// TIA Portal V21 export
// export: Created 2026-11-22T02:34:22.6112688Z, ExportSetting WithDefaults, DisplayName Totally Integrated Automation Portal, DisplayVersion V21 Update 3, DisplayName STEP 7 Professional, DisplayVersion V21 Update 3, DisplayName STEP 7 Safety, DisplayVersion V21, DisplayName Tech WebApplication, DisplayVersion V21, DisplayName WinCC Basic/Comfort/Advanced, DisplayVersion V21 Update 3, DisplayName WinCC Unified, DisplayVersion V21 Update 3
TextList "TL_Value"  ListRange=Decimal
  TextListEntry   EntryType=Range, From=-100, To=-1, Text="Negative (-100..-1)"
  TextListEntry   EntryType=SingleValue, Text="Zero"
  TextListEntry   EntryType=Range, From=1, To=9, Text="One to nine"
  TextListEntry   EntryType=SingleValue, From=10, To=10, Text="Ten: Ünïcödé äöüß ÄÖÜ €"
  TextListEntry   EntryType=SingleValue, From=32000, To=32000, Text="Undefined value (default entry)"
